// Generated by voz_llm_plc_agent
// Target: Siemens TIA Portal V18 - SCL external source
// Review and compile before any download to physical hardware.

FUNCTION_BLOCK "PLC_PRG"
{ S7_Optimized_Access := 'TRUE' }
VERSION : 0.1
VAR_INPUT
   I_Emergency : Bool := FALSE;
   I_Lamp_Control : Bool := FALSE;
END_VAR
VAR_OUTPUT
   Q_Lamp : Bool := FALSE;
END_VAR
BEGIN
(* Salidas: contribucion automatica (secuencia/condiciones) y manual, con sus bloqueos *)
#Q_Lamp := (#I_Lamp_Control AND NOT #I_Emergency) AND NOT #I_Emergency;
END_FUNCTION_BLOCK

DATA_BLOCK "DB_PLC_PRG"
{ S7_Optimized_Access := 'TRUE' }
VERSION : 0.1
NON_RETAIN
"PLC_PRG"
BEGIN
END_DATA_BLOCK

ORGANIZATION_BLOCK "Main"
{ S7_Optimized_Access := 'TRUE' }
VERSION : 0.1
BEGIN
   "DB_PLC_PRG"(
      I_Emergency := "I_Emergency",
      I_Lamp_Control := "I_Lamp_Control",
      Q_Lamp => "Q_Lamp"
   );
END_ORGANIZATION_BLOCK
